# EPICS substitutions: niusb/niusbApp/Db/USB6008.substitutions
# The USB-6008: every record, by measComp's names (the 621x's where the meaning
# is the same). Macros: P, PORT, MAX_POINTS (from the entity); the templates at
# the image's /epics/support/niusb/db.
file "/epics/support/niusb/db/niusbDevice.template" { pattern {} {} }

file "/epics/support/niusb/db/niusb6008Ai.template"
{
pattern
{ N, ADDR }
{ 1, 0 }
{ 2, 1 }
{ 3, 2 }
{ 4, 3 }
{ 5, 4 }
{ 6, 5 }
{ 7, 6 }
{ 8, 7 }
}

file "/epics/support/niusb/db/niusbAo.template"
{
pattern
{ N, ADDR, DRVL, DRVH, LOPR, HOPR }
{ 1, 0, 0, 5, 0, 5 }
{ 2, 1, 0, 5, 0, 5 }
}

file "/epics/support/niusb/db/niusbBi.template"
{
pattern
{ N, LINE, MASK }
{ 1, 0, 0x1 }
{ 2, 1, 0x2 }
{ 3, 2, 0x4 }
{ 4, 3, 0x8 }
{ 5, 4, 0x10 }
{ 6, 5, 0x20 }
{ 7, 6, 0x40 }
{ 8, 7, 0x80 }
}

file "/epics/support/niusb/db/niusbBo.template"
{
pattern
{ N, LINE, MASK }
{ 1, 0, 0x1 }
{ 2, 1, 0x2 }
{ 3, 2, 0x4 }
{ 4, 3, 0x8 }
}

file "/epics/support/niusb/db/niusb6008WaveDig.template" { pattern {} {} }

file "/epics/support/niusb/db/niusbWaveDigN.template"
{
pattern
{ N, ADDR }
{ 1, 0 }
{ 2, 1 }
{ 3, 2 }
{ 4, 3 }
{ 5, 4 }
{ 6, 5 }
{ 7, 6 }
{ 8, 7 }
}
